TYPE "FRK_ModelImage"
VERSION : 0.1
   STRUCT
      "Catalog" {ExternalAccessible := 'False'; ExternalVisible := 'False'; ExternalWritable := 'False'} : "FRK_ModelCatalog";
      "RecordCount" {ExternalAccessible := 'False'; ExternalVisible := 'False'; ExternalWritable := 'False'} : Int;
      "Rows" {ExternalAccessible := 'False'; ExternalVisible := 'False'; ExternalWritable := 'False'} : Array[1..5] of "FRK_ConfigSlot";
   END_STRUCT;
END_TYPE
